Fanuc KAREL source: KB00076.KL

PROGRAM KB00076
%NOLOCKGROUP
VAR
  P1: POSITION
  P2: POSITION
  P3: POSITION
  RESULT: POSITION
BEGIN
  RESULT = FRAME(P1, P2, P3)
END KB00076
